(* Logix 5000 project; controller TFF vendor 1 type 14 code 107 rev 33.11; software revision 33.04 *)
// Mobius TFF

TASK HighPriority (periodic, rate 25 ms, priority 1, watchdog 2000 ms) : MainProgram   // High Priority Task
TASK MainTask (continuous, watchdog 500 ms) : Process, CCPSystem
TASK Task5ms (periodic, rate 5 ms, priority 10, watchdog 500 ms) : MainProgram5ms

MODULES
   Local : vendor 1 type 14 code 107 (Compact 0, rev 33.11)
      GATEWAY : ETHERNET-MODULE (Ethernet 10.20.60.222, rev 1.1, Output RPI 50 ms)
           GATEWAY:I   // Gateway data from hardware
           GATEWAY:O   // Gateway data from hardware
           GATEWAY:C   // Gateway data from hardware
      GWModbus : ETHERNET-MODULE (Ethernet 10.20.60.200, rev 1.1, Output RPI 50 ms)
           GWModbus:I.Data[56]   // R_PMC1 Unit
           GWModbus:I.Data[0]   // R_User Level
           GWModbus:I.Data[100]   // R_Warning Interface
           GWModbus:I.Data[101]   // R_Warning Interface
           GWModbus:I.Data[102]   // R_Warning Hardware
           GWModbus:I.Data[103]   // R_Warning Hardware
           GWModbus:I.Data[10]   // R_PMC1 Min limit
           GWModbus:I.Data[11]   // R_PMC1 Min limit
           GWModbus:I.Data[12]   // R_PMC1 Max limit
           GWModbus:I.Data[13]   // R_PMC1 Max limit
           GWModbus:I.Data[14]   // R_CalibStatus Status
           GWModbus:I.Data[15]   // R_CalibStatus Status
           GWModbus:I.Data[16]   // R_CalibStatus Unit
           GWModbus:I.Data[17]   // R_CalibStatus Unit
           GWModbus:I.Data[18]   // R_CalibStatus Value
           GWModbus:I.Data[19]   // R_CalibStatus Value
           GWModbus:I.Data[1]   // R_User Level
           GWModbus:I.Data[20]   // R_CalibLimits Offset Min
           GWModbus:I.Data[21]   // R_CalibLimits Offset Min
           GWModbus:I.Data[22]   // R_CalibLimits Offset Max
           GWModbus:I.Data[23]   // R_CalibLimits Offset Max
           GWModbus:I.Data[24]   // R_CalibLimits Slope Min
           GWModbus:I.Data[25]   // R_CalibLimits Slope Min
           GWModbus:I.Data[26]   // R_CalibLimits Slope Max
           GWModbus:I.Data[27]   // R_CalibLimits Slope Max
           GWModbus:I.Data[28]   // R_CalibValues Offset
           GWModbus:I.Data[29]   // R_CalibValues Offset
           GWModbus:I.Data[2]   // R_User N/A
           GWModbus:I.Data[30]   // R_CalibValues Slope
           GWModbus:I.Data[31]   // R_CalibValues Slope
           GWModbus:I.Data[32]   // R_CalibValues Temp
           GWModbus:I.Data[33]   // R_CalibValues Temp
           GWModbus:I.Data[34]   // R_CalibAct pH
           GWModbus:I.Data[35]   // R_CalibAct pH
           GWModbus:I.Data[36]   // R_CalibAct Elec
           GWModbus:I.Data[37]   // R_CalibAct Elec
           GWModbus:I.Data[38]   // R_CalibAct Temp
           GWModbus:I.Data[39]   // R_CalibAct Temp
           GWModbus:I.Data[3]   // R_User N/A
           GWModbus:I.Data[40]   // R_CalibAct NA
           GWModbus:I.Data[41]   // R_CalibAct NA
           GWModbus:I.Data[42]   // R_CalibTime Time
           GWModbus:I.Data[43]   // R_CalibTime Time
           GWModbus:I.Data[44]   // R_Warning Measurement
           GWModbus:I.Data[45]   // R_Warning Measurement
           GWModbus:I.Data[46]   // R_Warning Calibration
           GWModbus:I.Data[47]   // R_Warning Calibration
           GWModbus:I.Data[48]   // R_Warning Interface
           GWModbus:I.Data[49]   // R_Warning Interface
           GWModbus:I.Data[4]   // R_PMC1 Unit
           GWModbus:I.Data[50]   // R_Warning Hardware
           GWModbus:I.Data[51]   // R_Warning Hardware
           GWModbus:I.Data[52]   // R_User Level
           GWModbus:I.Data[53]   // R_User Level
           GWModbus:I.Data[54]   // R_User N/A
           GWModbus:I.Data[55]   // R_User N/A
           GWModbus:I.Data[57]   // R_PMC1 Unit
           GWModbus:I.Data[8]   // R_PMC1 Status
           GWModbus:I.Data[58]   // R_PMC1 Value
           GWModbus:I.Data[59]   // R_PMC1 Value
           GWModbus:I.Data[5]   // R_PMC1 Unit
           GWModbus:I.Data[60]   // R_PMC1 Status
           GWModbus:I.Data[61]   // R_PMC1 Status
           GWModbus:I.Data[62]   // R_PMC1 Min limit
           GWModbus:I.Data[63]   // R_PMC1 Min limit
           GWModbus:I.Data[64]   // R_PMC1 Max limit
           GWModbus:I.Data[65]   // R_PMC1 Max limit
           GWModbus:I.Data[66]   // R_CalibStatus Status
           GWModbus:I.Data[67]   // R_CalibStatus Status
           GWModbus:I.Data[68]   // R_CalibStatus Unit
           GWModbus:I.Data[69]   // R_CalibStatus Unit
           GWModbus:I.Data[6]   // R_PMC1 Value
           GWModbus:I.Data[70]   // R_CalibStatus Value
           GWModbus:I.Data[71]   // R_CalibStatus Value
           GWModbus:I.Data[72]   // R_CalibLimits Offset Min
           GWModbus:I.Data[73]   // R_CalibLimits Offset Min
           GWModbus:I.Data[74]   // R_CalibLimits Offset Max
           GWModbus:I.Data[75]   // R_CalibLimits Offset Max
           GWModbus:I.Data[76]   // R_CalibLimits Slope Min
           GWModbus:I.Data[77]   // R_CalibLimits Slope Min
           GWModbus:I.Data[78]   // R_CalibLimits Slope Max
           GWModbus:I.Data[79]   // R_CalibLimits Slope Max
           GWModbus:I.Data[7]   // R_PMC1 Value
           GWModbus:I.Data[80]   // R_CalibValues Offset
           GWModbus:I.Data[81]   // R_CalibValues Offset
           GWModbus:I.Data[82]   // R_CalibValues Slope
           GWModbus:I.Data[83]   // R_CalibValues Slope
           GWModbus:I.Data[84]   // R_CalibValues Temp
           GWModbus:I.Data[85]   // R_CalibValues Temp
           GWModbus:I.Data[86]   // R_CalibAct pH
           GWModbus:I.Data[87]   // R_CalibAct pH
           GWModbus:I.Data[88]   // R_CalibAct Elec
           GWModbus:I.Data[89]   // R_CalibAct Elec
           GWModbus:I.Data[9]   // R_PMC1 Status
           GWModbus:I.Data[90]   // R_CalibAct Temp
           GWModbus:I.Data[91]   // R_CalibAct Temp
           GWModbus:I.Data[92]   // R_CalibAct NA
           GWModbus:I.Data[93]   // R_CalibAct NA
           GWModbus:I.Data[94]   // R_CalibTime Time
           GWModbus:I.Data[95]   // R_CalibTime Time
           GWModbus:I.Data[96]   // R_Warning Measurement
           GWModbus:I.Data[97]   // R_Warning Measurement
           GWModbus:I.Data[98]   // R_Warning Calibration
           GWModbus:I.Data[99]   // R_Warning Calibration
           GWModbus:O.Data[12]   // W_CalibValue Temp
           GWModbus:O.Data[0]   // W_User Level
           GWModbus:O.Data[10]   // W_CalibValue Slope
           GWModbus:O.Data[11]   // W_CalibValue Slope
           GWModbus:O.Data[13]   // W_CalibValue Temp
           GWModbus:O.Data[24]   // W_SysTime Trigger
           GWModbus:O.Data[14]   // W_CalibProd Trigger
           GWModbus:O.Data[15]   // W_CalibProd Command
           GWModbus:O.Data[16]   // W_CalibProd Command
           GWModbus:O.Data[17]   // W_CalibProdVal Trigger
           GWModbus:O.Data[18]   // W_CalibProdVal Value
           GWModbus:O.Data[19]   // W_CalibProdVal Value
           GWModbus:O.Data[1]   // W_User Level
           GWModbus:O.Data[20]   // W_User Level
           GWModbus:O.Data[21]   // W_User Level
           GWModbus:O.Data[22]   // W_User Password
           GWModbus:O.Data[23]   // W_User Password
           GWModbus:O.Data[32]   // W_CalibValue Temp
           GWModbus:O.Data[25]   // W_SysTime Time
           GWModbus:O.Data[26]   // W_SysTime Time
           GWModbus:O.Data[27]   // W_CalibValue Trigger
           GWModbus:O.Data[28]   // W_CalibValue Offset
           GWModbus:O.Data[29]   // W_CalibValue Offset
           GWModbus:O.Data[2]   // W_User Password
           GWModbus:O.Data[30]   // W_CalibValue Slope
           GWModbus:O.Data[31]   // W_CalibValue Slope
           GWModbus:O.Data[33]   // W_CalibValue Temp
           GWModbus:O.Data[8]   // W_CalibValue Offset
           GWModbus:O.Data[34]   // W_CalibProd Trigger
           GWModbus:O.Data[35]   // W_CalibProd Command
           GWModbus:O.Data[36]   // W_CalibProd Command
           GWModbus:O.Data[37]   // W_CalibProdVal Trigger
           GWModbus:O.Data[38]   // W_CalibProdVal Value
           GWModbus:O.Data[39]   // W_CalibProdVal Value
           GWModbus:O.Data[3]   // W_User Password
           GWModbus:O.Data[4]   // W_SysTime Trigger
           GWModbus:O.Data[5]   // W_SysTime Time
           GWModbus:O.Data[6]   // W_SysTime Time
           GWModbus:O.Data[7]   // W_CalibValue Trigger
           GWModbus:O.Data[9]   // W_CalibValue Offset
      RACK_ACT350_WI101_200L : ETHERNET-MODULE (Ethernet 10.20.60.142, rev 1.1, Output RPI 50 ms)
      RACK_ACT350_WI101_500L : ETHERNET-MODULE (Ethernet 10.20.60.141, rev 1.1, Output RPI 50 ms)
      RACK_MURR_NODE0_SMART : ETHERNET-MODULE (Ethernet 10.20.60.131, rev 1.1, Output RPI 50 ms)
           RACK_MURR_NODE0_SMART:I   // Node 0 data from hardware
           RACK_MURR_NODE0_SMART:O.Data[0]   // MOM
           RACK_MURR_NODE0_SMART:O.Data[1]   // MOM
           RACK_MURR_NODE0_SMART:O.Data[2]   // MOM
           RACK_MURR_NODE0_SMART:O.Data[3]   // MOM
           RACK_MURR_NODE0_SMART:O.Data[4]   // MOM
           RACK_MURR_NODE0_SMART:O.Data[5]   // MOM
           RACK_MURR_NODE0_SMART:O.Data[6]   // Bus Control
           RACK_MURR_NODE0_SMART:O.Data[7]   // Bus Control
           RACK_MURR_NODE0_SMART:O   // Node 0 data from hardware
           RACK_MURR_NODE0_SMART:C   // Node 0 data from hardware
      RACK_MURR_NODE1_TFF20 : ETHERNET-MODULE (Ethernet 10.20.60.123, rev 1.1, Output RPI 5 ms)
           RACK_MURR_NODE1_TFF20:C   // Node 1 data from hardware
           RACK_MURR_NODE1_TFF20:I   // Node 1 data from hardware
           RACK_MURR_NODE1_TFF20:O   // Node 1 data from hardware
      RACK_MURR_NODE1_TFF40 : ETHERNET-MODULE (Ethernet 10.20.60.124, rev 1.1, Output RPI 5 ms)
           RACK_MURR_NODE1_TFF40:I   // Node 1 data from hardware
           RACK_MURR_NODE1_TFF40:O   // Node 1 data from hardware
           RACK_MURR_NODE1_TFF40:C   // Node 1 data from hardware
      RACK_MURR_NODE1_TFF80 : ETHERNET-MODULE (Ethernet 10.20.60.126, rev 1.1, Output RPI 5 ms)
           RACK_MURR_NODE1_TFF80:I   // Node 1 data from hardware
           RACK_MURR_NODE1_TFF80:O   // Node 1 data from hardware
           RACK_MURR_NODE1_TFF80:C   // Node 1 data from hardware
END_MODULES

TYPE AlarmAnalog :   // Analog Alarm UDT
STRUCT
   Override : BOOL;   // Alarm Override
   Disable : BOOL;   // Alarm Disabled
   LOLOAlarm : BOOL;   // LOLO Alarm Condition
   LOAlarm : BOOL;   // LO Alarm Condition
   HIAlarm : BOOL;   // HI Alarm Condition
   HIHIAlarm : BOOL;   // HIHI Alarm Condition
   LOLODisable : BOOL;   // LOLO Alarm Disable
   LODisable : BOOL;   // LO Alarm Disable
   HIDisable : BOOL;   // HI Alarm Disable
   HIHIDisable : BOOL;   // HIHI Alarm Disable
   LOLOAck : BOOL;   // LOLO Alarm Acknowledged
   LOAck : BOOL;   // LO Alarm Acknowledged
   HIAck : BOOL;   // HI Alarm Acknowledged
   HIHIAck : BOOL;   // HIHI Alarm Acknowledged
   HIHIEnable : BOOL;   // HIHI Alarm Always Enabled for Critical Safety Alarms
   FeedPumpEnable : BOOL;   // LOLO and LO Alarm conditionned on Feed Pump Enable
   TransferPumpEnable : BOOL;   // LOLO and LO Alarm conditionned on Transfer Pump Enable
   LOLOAlarmONS : BOOL;   // Saves last value of alarm
   LOAlarmONS : BOOL;   // Saves last value of alarm
   HIAlarmONS : BOOL;   // Saves last value of alarm
   HIHIAlarmONS : BOOL;   // Saves last value of alarm
   FeedPumpTag : DINT;   // Feed Pump Tag for Pump Enable function
   TransferPumpTag : DINT;   // Transfer Pump Tag for Pump Enable function
   Value : DINT;   // Alarm Value : 0= No Alarm. 1=Non-Critical. 2= Non-Critical Unacknowledged. 3=Critical. 4=Critical Unacknowledged.
   ValueHMI : DINT;   // Alarm Value for HMI: 0= No Alarm. 1=Non-Critical. 2= Non-Critical Unacknowledged. 3=Critical. 4=Critical Unacknowledged.
   LOLO : REAL;   // LOLO Alarm Set Point
   LO : REAL;   // LO Alarm Set Point
   HI : REAL;   // HI Alarm Set Point
   HIHI : REAL;   // HIHI Alarm Set Point
   PV : REAL;   // Process Variable Value
   LOLOTimer : TIMER;   // LOLO Alarm Timer
   LOLOTimerSP : DINT;   // LOLO Alarm Timer setpoint (sec)
   LOTimer : TIMER;   // LO Alarm Timer
   LOTimerSP : DINT;   // LO Alarm Timer setpoint (sec)
   HITimer : TIMER;   // HI Alarm Timer
   HITimerSP : DINT;   // HI Alarm Timer setpoint (sec)
   HIHITimer : TIMER;   // HIHI Alarm Timer
   HIHITimerSP : DINT;   // HIHI Alarm Timer setpoint (sec)
   EnableCfg : BOOL;   // Set to 1 to Configure \ Use Analog Alarm
END_STRUCT
END_TYPE

TYPE AlarmControl :   // Alarm Control UDT
STRUCT
   DESC : STRING25;   // Description
   EGU : STRING5;   // Unit
   InitAlarmconfig : BOOL;   // Initialize alarms config if the command is set from the HMI
   AlarmAck : BOOL;   // Alarm Acknowledge Flag
   AlarmHigh : BOOL;   // Critical Alarm Condition
   AlarmLow : BOOL;   // Non-Critical Alarm Condition
   AlarmHighUnack : BOOL;   // Critical Unacknowledged Alarm Condition
   AlarmLowUnack : BOOL;   // Non-Critical Unacknowledged Alarm Condition
   HighHMI : BOOL;   // Critical Alarm Condition (for HMI)
   LowHMI : BOOL;   // Non-Critical Alarm Condition (for HMI)
   HighUnackHMI : BOOL;   // Critical Unacknowledged Alarm Condition (for HMI)
   LowUnackHMI : BOOL;   // Non-Critical Unacknowledged Alarm Condition (for HMI)
   Horn : BOOL;   // Alarm Horn
   YellowLamp : BOOL;   // Non-Critical Alarm Indicator
   RedLamp : BOOL;   // Critical Alarm Indicator
   Current : BOOL;   // Current Alarm Status
   AckOutput : BOOL;   // Alarm Acknowledge Output
   FlashControl : BOOL;   // Flash Control
   LightingBannercfg : BOOL;   // Lighting Banner configuration (1= ON)
   EnableAllIn : BOOL;   // Enable All Alarms Input
   EnableAllOut : BOOL;   // Enable All Alarms Output
   DisableAllIn : BOOL;   // Disable All Alarms Input
   DisableAllOut : BOOL;   // Disable All Alarms Output
   NewAlarm : BOOL;   // True for 1 scan when new alarm is detected
   SilenceHorn : BOOL;   // Set true to Silence horn
   FlashTimer : TIMER;   // Flash Timer
   AckTimer : TIMER;   // Acknowledge Timer
   EnableAllTimer : TIMER;   // Enable All Alarms Timer
   DisableAllTimer : TIMER;   // Disable All Alarms Timer
   EnableAllAnaSigIn : BOOL;   // Enable All analog signal failure Alarms Input
   EnableAllAnaSigOut : BOOL;   // Enable All analog signal failure Alarms Output
   DisableAllAnaSigIn : BOOL;   // Disable All analog signal failure Alarms Input
   DisableAllAnaSigOut : BOOL;   // Disable All analog signal failure Alarms Output
   EnableAllAnaSigTimer : TIMER;   // Enable All analog signal failure Alarms Timer
   DisableAllAnaSigTimer : TIMER;   // Disable All analog signal failure Alarms Timer
   AlarmHighMem : BOOL;   // Critical Alarm Condition Mem
END_STRUCT
END_TYPE

TYPE AlarmDeviation :   // Deviation Alarm UDT
STRUCT
   Override : BOOL;   // Alarm Override
   Disable : BOOL;   // Alarm Disabled
   HIAlarm : BOOL;   // HI Deviation Alarm Condition
   HIHIAlarm : BOOL;   // HIHI Deviation Alarm Condition
   HIDisable : BOOL;   // HI Alarm Disable
   HIHIDisable : BOOL;   // HIHI Alarm Disable
   HIAck : BOOL;   // HI Alarm Acknowledged
   HIHIAck : BOOL;   // HIHI Alarm Acknowledged
   LOLOAlarmONS : BOOL;   // One shot when alarm occures
   HIAlarmONS : BOOL;   // One shot when alarm occures
   LOAlarmONS : BOOL;   // One shot when alarm occures
   HIHIAlarmONS : BOOL;   // One shot when alarm occures
   Value : DINT;   // Alarm Value
   ValueHMI : DINT;   // Alarm Value for HMI
   HI : REAL;   // HI Alarm Set Point
   HIHI : REAL;   // HIHI Alarm Set Point
   LOLOLim : REAL;   // LOLO Alarm Set Point (calculated)
   LOLim : REAL;   // LO Alarm Set Point (calculated)
   HILim : REAL;   // HI Alarm Set Point (calculated)
   HIHILim : REAL;   // HIHI Alarm Set Point (calculated)
   HITimer : TIMER;   // HI Alarm Timer
   HITimerSP : DINT;   // HI Alarm Timer setpoint (sec)
   HIHITimer : TIMER;   // HIHI Alarm Timer
   HIHITImerSP : DINT;   // HIHI Alarm Timer setpoint (sec)
   EnableCfg : BOOL;   // Set to enable alarm
END_STRUCT
END_TYPE

TYPE AnalogInput :   // Analog Input UDT
STRUCT
   TagName : STRING6;   // PID Tag Name
   TagDisplayName : STRING6;   // PID Tag Name
   OutofRange : BOOL;   // Out of Range
   FilterType : BOOL;   // Filter Type 0=LP, 1=Avg
   AveragingTotal : DINT;   // Averaging Filter Total
   Address : DINT;   // Input Address (RawAnalogInputArray)
   RawMin : DINT;   // Raw Minimum Range
   RawMax : DINT;   // Raw Maximum Range
   RawValue : DINT;   // Raw Value (Measuring value given by the I/O card)
   RawLowLimit : DINT;   // Raw Out of Range LO Limit
   RawHighLimit : DINT;   // Raw Out of Range HI Limit
   FilterUser : DINT;   // User Filter Value
   FilteredRaw : DINT;   // Raw Filtered Value
   FilterActual : REAL;   // Actual Filter Value
   ScaledMin : REAL;   // Scaled Minimum Range
   ScaledMax : REAL;   // Scaled Maximum Range
   CurrentValue : REAL;   // Current Value
   RangeMin : REAL;   // Scaled Minimum Range (Config Analog Points)
   RangeMax : REAL;   // Scaled Maximum Range (Config Analog Points)
   RangeMinSave : REAL;   // Scaled Minimum Range (previous)
   RangeMaxSave : REAL;   // Scaled Maximum Range (previous)
   RealCfg : BOOL;   // Set to 1 if real analog input is used. Set to 0 for soft input (derived data)
   EnableCfg : BOOL;   // Set to 1 to activate this Tag
   OverrideCfg : BOOL;   // Set to 1 to allow user to Overide alarm
   Desc : STRING25;   // Description
   EGU : STRING5;   // Unit
END_STRUCT
END_TYPE

TYPE AnalogOutput :   // Analog Output UDT
STRUCT
   Tag : STRING10;   // Tag name
   RawValue : DINT;   // Raw Value Send to I/O Card
   RawMin : DINT;   // Raw Min
   RawMax : DINT;   // Raw Max
   ScaledValue : REAL;   // Scaled Value
   ScaledMin : REAL;   // Scaled Minimum Range
   ScaledMax : REAL;   // Scaled Maximum Range
   EnableCfg : BOOL;   // Set to 1 to enable Analog Output
END_STRUCT
END_TYPE

TYPE ARC_pH :   // ARC pH Communication Structure
STRUCT
   SetCalibValues : BOOL;   // Set calibration values from HMI
   ActiveCalibration : BOOL;   // Current Active Calibration (0= Standrad, 1= Product)
   ActiveCalibrationSave : BOOL;   // Save state of Active Calibration
   AssignedCalibration : BOOL;   // Product Calibration is assigned
   ActiveInitial : BOOL;   // Initial Measurement of Product Calibration has been taken
   WarningSetCalib : BOOL;   // Verify/Set Calibration Data Warning from device
   ProductReadInitial : BOOL;   // Read command for the Product Calibration Initial Measurment
   ProductAssign : BOOL;   // Submit the Product Assign value command
   ProductAssignTime : DINT;   // Time of the last Product Assign
   ProductAssignONS : BOOL;   // ONS for Product Assignment
   R_CALIBSTATUS_Status : DINT;   // Calibration status from register 5318
   R_CALIBSTATUS_Unit : DINT;   // Calibration unit from register 5318
   R_CALIBSTATUS_Value : REAL;   // Calibration value from register 5318
   R_CALIBLIMITS_MinOffset : REAL;   // Calibration Minimum value for Offset from register 5480
   R_CALIBLIMITS_MaxOffset : REAL;   // Calibration Maximum value for Offset from register 5480
   R_CALIBLIMITS_MinSlope : REAL;   // Calibration Minimum value for Slope from register 5480
   R_CALIBLIMITS_MaxSlope : REAL;   // Calibration Maximum value for Slope from register 5480
   W_CALIBVALUES_Trigger : BOOL;   // Write to register 5448
   W_CALIBVALUES_Offset : REAL;   // Calibration offset to register 5448
   W_CALIBVALUES_Slope : REAL;   // Calibration slope to register 5448
   W_CALIBVALUES_Temp : REAL;   // Calibration temperature to register 5448
   R_CALIBVALUES_Offset : REAL;   // Calibration offset from register 5448
   R_CALIBVALUES_Slope : REAL;   // Calibration slope from register 5448
   R_CALIBVALUES_Temp : REAL;   // Calibration temperature from register 5448
   W_CALIBPROD_Trigger : BOOL;   // Write to register 5340
   W_CALIBPROD_Command : DINT;   // Product calibration command to register 5340
   W_CALIBPRODVAL_Trigger : BOOL;   // Write to register 5322
   W_CALIBPRODVAL_Value : REAL;   // Product calibration value to register 5322
   R_CALIBACTUAL_PH : REAL;   // pH at initial calibration from register 5560
   R_CALIBACTUAL_Voltage : REAL;   // Voltage at initial calibration from register 5560
   R_CALIBACTUAL_Temp : REAL;   // Temparature at initial calibration from register 5560
   R_CALIBACTUAL_NA : REAL;   // Unused from register 5560
   R_CALIBTIME_Time : DINT;   // Date Time of last calibration from register 5342 (UNIX)
   W_SYNCTIME_Trigger : BOOL;   // Write to register 8232
   W_SYNCTIME_Time : DINT;   // Time to register 8232 (UNIX)
   R_PMC1_Unit : DINT;   // Value unit from register 2090
   R_PMC1_Value : REAL;   // Value from register 2090
   R_PMC1_Status : DINT;   // Value Status from register 2090
   R_PMC1_Min : REAL;   // Value Minimum Limit from register 2090
   R_PMC1_Max : REAL;   // Value Maximum Limit from register 2090
   W_USER_Level : DINT;   // User Level to register 4288
   W_USER_Password : DINT;   // User Password to register 4288
   R_USER_Level : DINT;   // User Level from register 4288
   R_WARNING_Calib : DINT;   // Calibration warning from register 4736
END_STRUCT
END_TYPE

TYPE BagInflate :   // Inflate Bag
STRUCT
   cmd : BOOL;   // Command form HMI
   SP : REAL;   // Pressure Setpoint from HMI
   PV : REAL;   // Current Pressure
END_STRUCT
END_TYPE

TYPE CCPSystem :   // CCP System UDT
STRUCT
   Run : BOOL;   // Run Flag
   RunAuto : BOOL;   // Auto Run Flag
   Procedure : BOOL;   // Procedure Flag
   Complete : BOOL;   // Procedure Complete
   Download : BOOL;   // Manual Download
   Heartbeat : BOOL;   // CCPRuntime Heartbeat
   OperationDownloadFlag : BOOL;   // Legacy Tag. Not used by PLC
   OperationStartFlag : BOOL;   // Operation Start Flag
   Manual : BOOL;   // Recipe Pool Flag
   State : DINT;   // Machine State
   Language : DINT;   // Language Number
   ErrorPhase : DINT;   // Error in Phase #
   ErrorStep : DINT;   // Error in Step #
   Error : DINT;   // Error Description
   OperationNoInBatch : DINT;   // Legacy Tag. Not used by PLC
   EndPointer : DINT;   // End Operation Step Buffer Pointer
   Machine : STRING;   // Machine Name
   ProductID : STRING;   // Batch Product ID from Operation Header
   Description : STRING;   // Batch Description from Operation Header
   Created : STRING;   // Date and Time when the last operation has been downloaded in PLC
   Originator : STRING;   // Last saved by field from Operation Header
   Comment : STRING;   // Comment
   OperationName : STRING90;   // Name and path of last operation downloaded in PLC
   ConfigFile : STRING;   // Current configuration file used
   LastMod : STRING;   // Last Mod
   GradientBasis : STRING;   // Gradient Basis
   GradientVariable : STRING;   // Gradient Variable
   GradientSegments : STRING;   // Gradient Segments
   StateWatchDog : TIMER;   // If Downloading for longer than this time the state will reset to 0
   EventList : EventList;   // Event List Array
   BufferSteps : STRING25[251];   // Buffer Steps Array
   BufferEvents : STRING50[251];   // Buffer Events Array
   HETP_ON_OFF : BOOL;   // HETP (1 = Start , 0 = Stop)
   DefaultOnComplete : BOOL;   // At the end of recipe apply default flowpath (0 = Apply , 1 = Don't Apply)
END_STRUCT
END_TYPE

TYPE CCPSystem_Storage :
STRUCT
   Run : BOOL;   // Run Flag
   RunAuto : BOOL;   // Auto Run Flag
   Procedure : BOOL;   // Procedure Flag
   Complete : BOOL;   // Procedure Complete
   Download : BOOL;   // Manual Download
   Heartbeat : BOOL;   // CCPRuntime Heartbeat
   OperationDownloadFlag : BOOL;   // Legacy Tag. Not used by PLC
   OperationStartFlag : BOOL;   // Operation Start Flag
   TestAction : BOOL;   // Action Test Flag
   Manual : BOOL;   // Recipe Pool Flag
   State : DINT;   // Machine State
   Language : DINT;   // Language Number
   ErrorPhase : DINT;   // Error in Phase #
   ErrorStep : DINT;   // Error in Step #
   Error : DINT;   // Error Description
   OperationNoInBatch : DINT;   // Legacy Tag. Not used by PLC
   EndPointer : DINT;   // End Operation Step Buffer Pointer
   Machine : STRING;
   ProductID : STRING;
   Description : STRING;
   Created : STRING;
   Originator : STRING;
   Comment : STRING;
   OperationName : STRING90;
   ConfigFile : STRING;
   LastMod : STRING;
   GradientBasis : STRING;
   GradientVariable : STRING;
   GradientSegments : STRING;
   StateWatchDog : TIMER;   // If Downloading for longer than this time the state will reset to 0
END_STRUCT
END_TYPE

TYPE ChartMark :   // Chart Mark UDT
STRUCT
   In : BOOL;   // Chart Mark In
   Out : BOOL;   // Chart Mark Out
END_STRUCT
END_TYPE

TYPE Concentration :   // Concentration UDT
STRUCT
   VCF : REAL;   // Volume Concentration Factor
   CB : REAL;   // Protein Concentration
   Conc_Init : REAL;   // Initial Protein Concentration SP
   Conc_Final : REAL;   // Final Protein Concentration SP
   Conc_Final_Volume : REAL;   // Final Concentration Volume SP
   Final_Conc_Volume_Reached : BOOL;   // Final Concentration Volume Reached
   Final_Conc_Protein_Reached : BOOL;   // Final Protein Concentration Reached
   LogConcIn : BOOL;   // Log Concentration Input
   LogConcOut : BOOL;   // Log Concentration Output
   LogConcTimer : TIMER;   // Log Concentation Timer
END_STRUCT
END_TYPE

TYPE Configuration :   // Configuration UDT
STRUCT
   Reset : BOOL;   // Activate Reset Loop Configuration
   IndexA0 : DINT;   // Index AnalogOutput
   IndexAP : DINT;   // Index AnalogPoint
   IndexDP : DINT;   // Index DigitalPoint
   IndexDr : DINT;   // Index Drive
   IndeXValve : DINT;   // Index Valve
   IndexReset : DINT;   // Index Reset
   IndexCL : DINT;   // Index Control Loop
   IndexFlowpath : DINT;   // Index Flowpath
   IndexIOMod : DINT;   // Index IO Module
END_STRUCT
END_TYPE

TYPE ControlLoop :   // Control Loop UDT
STRUCT
   Tag : STRING5;   // Tag Name
   Desc : STRING25;   // Description
   LoopCfg : BOOL;   // Set to 1 to use this loop
   ManualEGU : STRING5;   // Unit of Manual Control Mode
   AutoEGU : STRING5;   // Unit of Auto Control Mode
   Auto1EGU : STRING5;   // Unit of Auto Control Mode 1
   Auto2EGU : STRING5;   // Unit of Auto Control Mode 2
   Auto3EGU : STRING5;   // Unit of Auto Control Mode 3
   Interlock : BOOL;   // Loop Interlock
   Enable : BOOL;   // Loop Enabled
   Manual : BOOL;   // Control Mode 0=Auto, 1=Manual
   Stable : BOOL;   // Loop Stable
   DBOK : BOOL;   // Control Within Deadband
   Status : INT;   // Status
   Auto1 : BOOL;   // Auto Control Mode 1
   Auto2 : BOOL;   // Auto Control Mode 2
   Auto3 : BOOL;   // Auto Control Mode 3
   Auto4 : BOOL;   // Auto Control Mode 4
   StepUp : BOOL;   // Increment CV
   StepDown : BOOL;   // Decrement CV
   RampEnable : BOOL;   // Ramp Enable
   RampUp : BOOL;   // Ramping UP
   RampDown : BOOL;   // Ramping Down
   RampStatus : BOOL;   // Ramping Status
   RampAutoOSR : BOOL;   // Auto Ramp One-Shot
   RampManualOSR : BOOL;   // Manual Ramp One-Shot
   PIDEnable : BOOL;   // PID Enabled
   ManualOSR : BOOL;   // Manual Mode One-Shot
   Auto1OSR : BOOL;   // Control Mode 1 One-Shot
   Auto2OSR : BOOL;   // Control Mode 2 One-Shot
   Auto3OSR : BOOL;   // Control Mode 3 One-Shot
   Auto4OSR : BOOL;   // Control Mode 4 One-Shot
   StepIncrement : DINT;   // Step Increment/Decrement Value
   CycleTime : DINT;   // Cycle Time (for modulating output)
   PV : REAL;   // Process Variable
   PVAuto1 : REAL;   // Process Variable for Control Mode Auto 1
   PVAuto2 : REAL;   // Process Variable for Control Mode Auto 2
   PVAuto3 : REAL;   // Process Variable for Control Mode Auto 3
   PVAuto4 : REAL;   // Process Variable for Control Mode Auto 4
   CV : REAL;   // Control Value
   SPAuto : REAL;   // Auto Set Point
   SPAutoSave : REAL;   // Auto Set Point (previous)
   SPAuto1 : REAL;   // Auto Set Point Mode 1
   SPAuto2 : REAL;   // Auto Set Point Mode 2
   SPAuto3 : REAL;   // Auto Set Point Mode 3
   SPAuto4 : REAL;   // Auto Set Point Mode 4
   SPManual : REAL;   // Manual Set Point
   SPManualSave : REAL;   // Manual Set Point (previous)
   RangeMin : REAL;   // Min EGU Range
   RangeMax : REAL;   // Max EGU Range
   SPRangeMin : REAL;   // Set Point Min EGU Range
   SPRangeMax : REAL;   // Set Point Max EGU Range
   RampRate : REAL;   // Ramp Rate
   RampRateSave : REAL;   // Ramp Rate (previous)
   RampStart : REAL;   // Ramp Start Value
   Deadband : REAL;   // Deadband
   DBLO : REAL;   // Low Deadband Value
   DBHI : REAL;   // High Deadband Value
   RampTimer : TIMER;   // Ramp Timer
   StableTimer : TIMER;   // Loop Stable Timer
   StableTime : DINT;   // Loop Stable Time setpoint (sec)
   PIDTimer : TIMER;   // PID Timer
   CycleTimer : TIMER;   // Cycle Timer (for modulating output)
   PID : PID;   // PID Instruction Data
   KP : REAL[3];   // Loop Gain from HMI
   KI : REAL[3];   // Loop Reset from HMI
   KD : REAL[3];   // Loop Rate from HMI
   DB : REAL[3];   // Loop Deadband from HMI
   On : BOOL;   // Turns all controll On
   DisOSR : BOOL;   // One Shot DisOSR
   OutputOn_OSR : BOOL;   // One Shot OutputOn_OSR
   OutputOff_OSR : BOOL;   // One Shot OutputOff_OSR
   DigitalOutput : BOOL;   // Output from loop in for descrete control
   RampCfg : BOOL;   // Set to 1 to Enable Ramp Option
   Auto1Cfg : BOOL;   // Set to 1 to use Auto 1 option
   Auto2Cfg : BOOL;   // Set to 1 to use Auto 2 option
   Auto3Cfg : BOOL;   // Set to 1 to use Auto 3 option
   Auto4Cfg : BOOL;   // Set to 1 to use Auto 4 option
   Auto1PVCfg : DINT;   // Set to Analog Point Number
   Auto2PVCfg : DINT;   // Set to Analog Point Number
   Auto3PVCfg : DINT;   // Set to Analog Point Number
   Auto4PVCfg : DINT;   // Set to Analog Point Number
   Auto1RangeMax : REAL;   // Set Point EGU Range Max
   Auto2RangeMax : REAL;   // Set Point EGU Range Max
   Auto3RangeMax : REAL;   // Set Point EGU Range Max
   Auto4RangeMax : REAL;   // Set Point EGU Range Max
   AutoSwitchEnable : BOOL;   // Set to 1 to allow loop to switch from auto1 to auto 2
   OutputAddress : INT;   // Set to analog output to use for this loop
   LoopStatus : INT;   // Loop Mode Status for HMI
END_STRUCT
END_TYPE

TYPE CriteriaFlag :   // Criteria Flag UDT
STRUCT
   Flag1 : BOOL;   // Criteria Flag 1 (1=ON , 0=OFF)
   Flag2 : BOOL;   // Criteria Flag 2 (1=ON , 0=OFF)
   Flag3 : BOOL;   // Criteria Flag 3 (1=ON , 0=OFF)
   Flag4 : BOOL;   // Criteria Flag 4 (1=ON , 0=OFF)
   Flag5 : BOOL;   // Criteria Flag 5 (1=ON , 0=OFF)
END_STRUCT
END_TYPE

TYPE CVTune :   // Control Valve Tuning Data Type
STRUCT
   ClosedRaw : REAL;   // Captured Raw Value When Valve is Closed
   OpenRaw : REAL;   // Captured Raw Value When Valve is Open
   MinOutput : REAL;   // Minimum output for tuning adjustment for valve
   MaxOutput : REAL;   // Maximum output for tuning adjustment for valve
   MinTimer : TIMER;   // Timer to capture closed raw value
   MaxTimer : TIMER;   // Timer to capture open raw value
   OSR : INT;   // One shot bits
   Activate : BOOL;   // Activate tuning function
   Enable : BOOL;   // Tuning routine is enabled
END_STRUCT
END_TYPE

TYPE DerivedData :   // DerivedData UDT
STRUCT
   HOLDUP : REAL;   // Holdup Volume
   FI101Q : REAL;   // Qmax Factor for FI101
   FI201Q : REAL;   // Qmax Factor for FI201
   FI401Q : REAL;   // Qmax Factor for FI401
   FI101K : REAL;   // K Factor for FI101
   FI201K : REAL;   // K Factor for FI201
   FI401K : REAL;   // K Factor for FI401
END_STRUCT
END_TYPE

TYPE Diafiltration :   // Diafiltration UDT
STRUCT
   Diaf_Volume : REAL;   // Diafiltration Volume
   Diaf_Init : REAL;   // Initial Diafiltration Volume SP
   Diaf_Final_Volume : REAL;   // Final Diafiltration Volume SP
   Snap : BOOL;   // Level Snapshot
   Final_Diaf_Volum_Reached : BOOL;   // Final Diafiltration Volume Reached
   Diaf_Snap_Value : REAL;   // Volume value snapped
   LogDiafIn : BOOL;   // Log Diafiltration Input
   LogDiafOut : BOOL;   // Log Diafiltration Output
   LogDiafTimer : TIMER;   // Log Diafiltration Timer
END_STRUCT
END_TYPE

TYPE DigitalPoint :   // Digital Point UDT
STRUCT
   Tag : STRING10;   // PID Tag to be Used for Display
   Desc : STRING25;   // Description to be Used for Display
   CurrentValue : BOOL;   // Current value of Tag
   AlarmCurrentValue : BOOL;   // Displays state of processed alarm input.
   AlarmAck : BOOL;   // Alarm Acknowledged
   Alarm : BOOL;   // Alarm
   Override : BOOL;   // Alarm Override
   Mimic : INT;   // Set color on HMI digital point mimic
   SoftInput : BOOL;   // Used as current value when RealInputCfg is set to 0
   Condition1 : BOOL;   // Enable Condition 1 Must be True to Enable alarm condition
   Condition2 : BOOL;   // Enable Condition 2 Must be True to Enable alarm condition
   Cond1Text : STRING;   // Condtion 1 Text
   Cond2Text : STRING;   // Condition 2 text
   DelayTimer : TIMER;   // Alarm Timer
   DelayTimerSP : DINT;   // Alarm Timer setpoint (sec)
   Priority : BOOL;   // Alarm Priority 0=Low, 1=High
   EnableCfg : BOOL;   // Set to True to configure point on system
   ActiveStateCFg : BOOL;   // Set to 0 to invert incomming state
   RealInputCfg : BOOL;   // Set to 1 to Use Hardwired Input. Set to 0 to disable Hardwired and use software condition
   InputAddressCfg : DINT;   // Set to address of hardwared input to be used on alarm
   AlarmCfg : BOOL;   // Set to 1 to Use alarm on this point
   AlarmStateCfg : BOOL;   // Set to 1 to alarm on a 0 to 1 transition. Set to zero to alarm on a 1 to 0 transition
   OverrideCfg : BOOL;   // set to 1 to allow user to Override alarm
   PriorityCfg : BOOL;   // Set to 1 to allow user to set Priority and Enable
   Cond1Cfg : BOOL;   // Set to 1 to Enable Condition
   Cond2Cfg : BOOL;   // Set to 1 to Enable Condition
   FlashingInputCfg : BOOL;   // Set to 1 for Heartbeat Style Inputs
   AlarmONS : BOOL;   // One shot when alarm occurs
END_STRUCT
END_TYPE

TYPE Drive :   // Pump Control UDT
STRUCT
   TagName : STRING10;   // Drive tag name
   Desc : STRING25;   // Drive Description
   Mode : BOOL;   // Control Mode
   ManualCommand : BOOL;   // Manual Command
   AutoCommand : BOOL;   // Auto Command
   RunCommand : BOOL;   // Run Command
   RunStatus : BOOL;   // Running Status
   RunInterlock : BOOL;   // Run Interlock
   RunInput : BOOL;   // Run Digital Input 0=No, 1=Yes
   OutputAddress : DINT;   // Run Command Output Address
   InputAddress : DINT;   // Running Input Address
   InterlockTimer : TIMER;   // Interlock Delay Timer
   RunOns : BOOL;   // Run one shot
   StopOns : BOOL;   // Stop One shot
   RunRequest : BOOL;   // Run request for auto or man mode
   Interlocked : BOOL;   // Drive is commanded to run but currently stopped by interlock
   EnableCfg : BOOL;   // Set to enable Drive
   ReverseCfg : BOOL;   // Set to enable reverse control
   Direction : BOOL;   // 0 = forward. 1 = reverse
   DirectionAddress : DINT;   // Direction Output Address
   DriveStatus : INT;   // Drive Status
   DriveLoopStatus : INT;   // Drive Loop Status
   DriveAlarmStatus : INT;   // Drive Alarm Status
   ValidFlowpath : BOOL;   // Valid flowpath flag
END_STRUCT
END_TYPE

TYPE EventList :
STRUCT
   Event : DINT[1000];   // Event List Array
   Value : REAL[1000];   // Value Array
   PreRunValue : REAL[1000];   // Pre Run Value
END_STRUCT
END_TYPE

TYPE Exchange_OUT :   // Exchange Output UDT
STRUCT
   AO01 : REAL;   // Exchange AO#1
   AO02 : REAL;   // Exchange AO#2
   AO03 : REAL;   // Exchange AO#3
   AO04 : REAL;   // Exchange AO#4
   DO01 : BOOL;   // Exchange DO#1
   DO02 : BOOL;   // Exchange DO#2
   DO03 : BOOL;   // Exchange DO#3
   DO04 : BOOL;   // Exchange DO#4
   DO05 : BOOL;   // Exchange DO#5
   DO06 : BOOL;   // Exchange DO#6
   DO07 : BOOL;   // Exchange DO#7
   DO08 : BOOL;   // Exchange DO#8
END_STRUCT
END_TYPE

TYPE FactorySettings :   // Factory Settings
STRUCT
   ProductName : STRING90;   // Product Name
   SerialNumber : STRING90;   // Serial Number
   ComputerName : STRING90;   // Computer Name
   ComputerDesc : STRING90;   // Computer Description
   DateFormat : STRING90;   // Date Format
   FlagUK : BOOL;   // Use UK Flag instead of US
   PCV101ClosedSP : REAL;   // PCV101 Closed SP
   PCV201ClosedSP : REAL;   // PCV201 Closed SP
   TCUDisableSP : REAL;   // TCU Disable SP
   BagInflateSP : REAL;   // Bag Inflate SP
END_STRUCT
END_TYPE

TYPE FaultRecordType :   // Fault Record Type UDT
STRUCT
   TimeLow : DINT;   // Lower 32 bits of the fault timestamp value
   TimeHigh : DINT;   // Upperer 32 bits of the fault timestamp value
   RecType : INT;   // Fault Type
   Code : INT;   // Unique code for the fault
   Info : DINT[8];   // Fault specific information
END_STRUCT
END_TYPE

TYPE FlowPath :   // Flow Path UDT
STRUCT
   Command : BOOL;   // Flow Path Command
   Status : BOOL;   // Flow Path Status
   Truth1 : DINT;   // Truth Table 1 (Valves 1-32)
   Truth2 : DINT;   // Truth Table 2 (Valves 33-64)
   Truth3 : DINT;   // Truth Table 3 (Valves 65-96)
   Truth4 : DINT;   // Truth Table 4 (Valves 97-128)
   Mask1 : DINT;   // Mask 1 (Valves 1-32)
   Mask2 : DINT;   // Mask 2 (Valves 33-64)
   Mask3 : DINT;   // Mask 3 (Valves 65-96)
   Mask4 : DINT;   // Mask 4 (Valves 97-128)
   Desc : STRING;   // Flow Path Description
END_STRUCT
END_TYPE

TYPE FlowPathControl :   // Flow Path Control UDT
STRUCT
   Flag : BOOL;   // Flow Path Command Flag
   Valve1 : DINT;   // Valve Control 1 (Valves 1-32)
   Valve2 : DINT;   // Valve Control 2 (Valves 33-64)
   Valve3 : DINT;   // Valve Control 3 (Valves 65-96)
   Valve4 : DINT;   // Valve Control 4 (Valves 97-128)
   MaxFlowPath : DINT;   // Maximum Number of Flow Paths
   Status : DINT;   // Flow Path Status
   StatusHMI : DINT;   // Flow Path Status for HMI
   Save : BOOL;   // Set to 1 to save Flowpath
   Restore : BOOL;   // Set to 1 to restore flowpath
   SaveOns : BOOL;   // one shot after save
   FlowpathEnable : BOOL[64];   // Enable Flowpath
   SaveStored : BOOL;   // Save the save cmd
   HoldOns : BOOL;   // one shot after hold
END_STRUCT
END_TYPE

TYPE FlowPathSetup :   // Flowpath Setup UDT
STRUCT
   Apply : BOOL;   // Apply Flow Path
   Number : DINT;   // Flow Path Number
   Prev : DINT;   // Previous Flow Path Number
   Mask_View : BOOL;   // View the Mask of selected Flowpath
   Mask_Save : BOOL;   // Save the Mask of selected Flowpath
   Truth_View : BOOL;   // View the Truth of selected Flowpath
   Truth_Save : BOOL;   // Save the Truth of selected Flowpath
   OpenAllValve : BOOL;   // Set the Flowpath 61 to Open All Valves
   CloseAllValve : BOOL;   // Set the Flowpath 62 to Close All Valves
END_STRUCT
END_TYPE

TYPE Gateway :   // Gateway UDT
STRUCT
   Inhibition : DINT;   // Inhibit \ Uninhibit Gateway Module
   Input : DINT[64];   // Swaped Data from Gateway
   Output : DINT[124];   // Swaped Data to Gateway
   RecipeAction_Digital : DINT[2];   // Data Send by PLC to Gateway (send from skid to customer) used as digital recipe action
   RecipeAction_Analog : REAL[20];   // Data Send by PLC to Gateway (send from skid to customer) used as analog recipe action
   RecipeCriteria_Digital : DINT[2];   // Data Read from the Gateway (receive from customer to skid) used as digital recipe criteria
   RecipeCriteria_Analog : REAL[20];   // Data Read from the Gateway (receive from customer to skid) used as analog recipe
   Watchdog_Heartbeat : BOOL;   // Gateway communication heartbeat
   Watchdog_Heartbeat_Timer : FBD_TIMER;   // Gateway communication heartbeat timer
   Watchdog_In_Ext : INT;   // Status data read by PLC (used to calculate customer watchdog)
   Watchdog_In_Skid : INT;   // Status data read by PLC (used to calculate skid watchdog)
   Watchdog_Out_Ext : INT;   // Status data send by PLC (used to calculate customer watchdog)
   Watchdog_Out_Skid : INT;   // Status data send by PLC (used to calculate skid watchdog)
   Index : DINT;   // Index
   Index2 : DINT;   // Index 2
END_STRUCT
END_TYPE

TYPE IO_Station :   // Station State UDT
STRUCT
   Node_Comm_Status_value : INT;   // Node Communication Status Value (get from status of hardware card)
   Node_Comm_Status : BOOL;   // Node Communication Status (0=Defect , 1=OK)
   Node_Internal_Defect_Status_value : INT;   // Node Internal Defect Status Value (at least one defect on the node : branch, slot, channel)
   Node_Internal_Defect_Status : BOOL;   // Node Internal Defect Status (0=Defect , 1=OK)
   Inhibition : DINT;   // Inhibit \ Uninhibit Station Module
   MOM_Mod_Config : BOOL[32];   // Activate \ Deactivate I/O Module (1 = Deactivate)
   MOM_Status : INT;   // Machine Option Management Status
   MOM_Restart : BOOL;   // 1 = Switch Off Voltage on modules , 0 = Restart the modules
   MOM_Enable_Config : BOOL;   // Enable modules configuration (avoid overwrite by options during the configuration)
END_STRUCT
END_TYPE

TYPE LinearGradient :   // Linear Gradient UDT
STRUCT
   Enable : BOOL;   // Linear Gradient Enable
   Hold : BOOL;   // Gradient Hold
   Segments : DINT;   // Number of Segments
   Variable : DINT;   // Gradient Variable (1=Time, 2=CVs, 3=Volume)
   Basis : DINT;   // Basis (1=Percent, 2=Conductivity)
   Segment : DINT;   // Current Segment
   State : DINT;   // Sets state of control : 0 = Disabled 1 = Running 2 = Paused
   Input : REAL;   // Input Value
   Result : REAL;   // Result
   X2 : REAL;   // Current Segment Duration
   Y1 : REAL;   // Current Start Value
   Y2 : REAL;   // Current End Value
   X : REAL[21];   // Gradient X Values (Durations)
   Y : REAL[21];   // Gradient Y Values (Set Points)
END_STRUCT
END_TYPE

TYPE LoggedValue :   // Logged Value UDT
STRUCT
   Value : REAL[8];   // Value to be logged in Audit Trail (used in Event section of configuration file)
END_STRUCT
END_TYPE

TYPE Membrane_Data :   // Membrane Data UDT
STRUCT
   Flux : REAL;   // Membrane Flux
   Area : REAL;   // Membrane Area SP
   Density : REAL;   // Density
   NWP_TCF : REAL;   // NWP Temperature correction factor
   NWP_TCF_Temp : INT;   // Temp. Temperature used in NWP calculation (INT)
   NWP_TCF_Lookup_25 : REAL[53];   // Lookup table for TCF
   AlarmStatus : INT;   // Alarm Status ( 0 = No Alarm , 1 = Non Critical Alarm , 2 = Critical Alarm )
END_STRUCT
END_TYPE

TYPE Memory_Data :   // This UDT is for putting the memory information returned by the Controller
STRUCT
   Reading_Request : BOOL;   // Request of Memory data reading
   Free_Mem_IO : DINT;   // Controler data: Free I/O Memory
   Free_Mem_DT : DINT;   // Controler data: Free Data & Logic Memory
   Free_Mem_Gen : DINT;   // Controler 1756-L55M16 only: Free Expansion Memory
   Free_Memory : DINT;   // Controler data: Total Free Memory (addition)
   Total_Mem_IO : DINT;   // Controler data: Total I/O Memory
   Total_Mem_DT : DINT;   // Controler data: Total Data & Logic Memory
   Total_Mem_Gen : DINT;   // Controler 1756-L55M16 only: Total Expansion Memory
   Total_Memory : DINT;   // Controler data: Total Memory (addition)
   Biggest_Gen_Mem_Size_Ava : DINT;   // Controler 1756-L55M16 only: Additionnal Expansion Memory
   Biggest_IO_Mem_Size_Ava : DINT;   // Controler 1756-L55M16 only: Largest contiguous block of Additionnal free Expansion Memory
   Biggest_DT_Mem_Size_Ava : DINT;   // Controler dsata: Largest contiguous block of Additionnal free Expansion Memory
   Total_Mem_DT_Real : REAL;   // Controler data: Total Data & Logic Memory
   Free_Mem_DT_Real : REAL;   // Controler data: Free Data & Logic Memory
   Used_Mem_DT_Real : REAL;   // Controler data: Used Data & Logic Memory
   Percentage_Used_DT : REAL;   // Controler data: Percentage of used Data & Logic Memory
END_STRUCT
END_TYPE

TYPE Mixer :
STRUCT
   Enable : BOOL;   // Enable Mixer Control Loop
   Mode : BOOL;   // Control Mode 0=Level, 1=Speed
   ModeONS : BOOL;   // Manual Mode One-Shot
   SPManual : REAL;   // Manual Speed Set Point
   SPAutoMin : REAL;   // Auto Max Speed Set Point
   SPAutoMax : REAL;   // Auto Min Speed Set Point
   LevelMin : REAL;   // Minimum Level
   LevelMax : REAL;   // Maximum Level
   CV : REAL;   // Control Value
   Alarm_Reset_Cmd : BOOL;   // Alarm Reset Command
   Alarm_Reset_Cmd_Timer : TIMER;   // Alarm Reset Command Timer
END_STRUCT
END_TYPE

TYPE OperatingTime :   // Operating Time Exceeded Control
STRUCT
   DayMax : REAL;   // Setpoint for Alarm Operating Time Exceeded
   HMICtrl : BOOL;   // Control Tag Reset on launch Workspace
   TimerCtrl : TIMER;   // Timer for set tag HMICtrl
   CountPre : DINT;   // Setpoint for Alarm in sec
   Counter : DINT;   // Second Counter for Alarm
END_STRUCT
END_TYPE

TYPE Operation :   // Operation UDT
STRUCT
   Step : DINT;   // Step Number
   Criteria1 : DINT;   // Criteria 1 Code
   Criteria1Operator : DINT;   // Criteria 1 Operator
   Boolean : DINT;   // Boolean
   Criteria2 : DINT;   // Criteria 2 Code
   Criteria2Operator : DINT;   // Criteria 2 Operator
   Action : DINT;   // Action Code
   Label : DINT;   // Label
   Criteria1Value : REAL;   // Criteria 1 Value
   Criteria2Value : REAL;   // Criteria 2 Value
   ActionValue : REAL;   // Action Value
END_STRUCT
END_TYPE

TYPE Options :   // Options UDT
STRUCT
   CCP_Report : BOOL;   // CCP Report
   InletFeed : BOOL;   // Feed Pump inlet
   InletFeed_Dis : BOOL;   // Feed Pump inlet Disabled
   FeedTank : BOOL;   // Feed Tank
   TransferFlow : BOOL;   // Transfer Flowmeter
   TankPH : BOOL;   // Tank pH Sensor
   TankCond : BOOL;   // Tank Conductivity Sensor
   FiltrateNoInstrum : BOOL;   // No Filtrate Instrument
   FiltrateNoInstrum_Dis : BOOL;   // No Filtrate Instrument Disabled
   FiltrateCondPH : BOOL;   // Filtrate Conductivity and PH
   FiltrateCondPHUV : BOOL;   // Filtrate Conductivity pH and UV
   FiltrateUltrasonicFlow : BOOL;   // Ultrasonic Filtrate Flowmeter instead of Magnetic
   FiltrateMagneticFlow : BOOL;   // Magnetic Filtrate Flowmeter instead of Ultrasonic
   SingleUsePH : BOOL;   // Single Use pH Sensor on Modbus Gateway
   External_IO : BOOL;   // External IO
   Gateway : BOOL;   // Gateway Anybus
   TFF80 : BOOL;   // TFF 80 Clamshell Installed
   TFF40 : BOOL;   // TFF 40 Clamshell Installed
   TFF20 : BOOL;   // TFF 20 Clamshell Installed
END_STRUCT
END_TYPE

TYPE PCV :
STRUCT
   SP : REAL;
   PV : REAL;
   ERREUR : REAL;
   CV : REAL;
   KP : REAL;
   KI : REAL;
   TP : REAL;
   TI : REAL;
   ACCU_TI : REAL;
   OpenRawValue : REAL;
   ClosedRawValue : REAL;
   RESET : BOOL;
END_STRUCT
END_TYPE

TYPE PCV_Calib :   // PCV Position Calibration
STRUCT
   Activate : BOOL;   // Calibration Command from HMI
   Enable : BOOL;   // PCV Calibration function enabled
   OSR : INT;   // One Shot bits
   Open_SP_Target : REAL;   // Open setpoint of PCV to achieve
   Close_SP_Target : REAL;   // Close setpoint of PCV to achieve
   Open_Timer : TIMER;   // Timer before save the raw value
   Close_Timer : TIMER;   // Timer before save the raw value
END_STRUCT
END_TYPE

TYPE PCV_Control :   // PCV Control UDT
STRUCT
   FullOpen : BOOL;   // fully open the valve without ramp
   FullOpenSP : REAL;   // target value of the valve opening
   FullOpenResetTimer : TIMER;   // Timer to reset full open command
   FullClose : BOOL;   // fully close the valve without ramp
   FullCloseSP : REAL;   // target value of the valve closing
   FullCloseResetTimer : TIMER;   // Timer to reset full close command
   ClosedStatusSP : REAL;   // Closed Status Setpoint
   ClosedStatus : BOOL;   // Closed Status
   CloseInterlocked : BOOL;   // Close Interlocked status for prohibit Manual Action on MHI
END_STRUCT
END_TYPE

TYPE Phases :   // Phase Control UDT
STRUCT
   Run : BOOL;   // Phase Run
   RunOSR : BOOL;   // Phase Run One-Shot
   Stop : BOOL;   // Phase Stop
   Hold : BOOL;   // Phase Hold
   Pause : BOOL;   // Phase Pause
   PauseOVR : BOOL;   // Pause Override
   Jump : BOOL;   // Phase Jump
   JumpPLC : BOOL;   // Phase Jump PLC
   Branch : BOOL;   // Branch Flag
   State : DINT;   // Phase State
   PendingStep : DINT;   // Pending Step Number
   JumpStep : DINT;   // Jump Step Number
   StartStep : DINT;   // Starting Step Number
   Crit1MetTime : DINT;   // Criteria 1 Met Timer
   NextStep : DINT;   // Next Step
   TotalSteps : DINT;   // Total Steps in Phase
   Label : DINT;   // Branch Label
   ActualStep : DINT;   // Actual Step
END_STRUCT
END_TYPE

TYPE PhaseTotalizer :   // Phase Totalizer UDT
STRUCT
   Enable : BOOL;   // Enable Totalizer
   PhaseEnable : BOOL;   // Enable Phase Totalizer
   StepEnable : BOOL;   // Enable Step Totalizer
   PauseEnable : BOOL;   // Enable Pause Totalizer
   UserEnable : BOOL;   // Enable User Totalizer
   ProcedureEnable : BOOL;   // Enable Procedure Totalizer
   PhaseReset : BOOL;   // Reset Phase Totalizer
   StepReset : BOOL;   // Reset Step Totalizer
   PauseReset : BOOL;   // Reset Pause Totalizer
   UserReset : BOOL;   // Reset User Totalizer
   PV : REAL;   // Totalizer Process Variable
   Phase : REAL;   // Phase Totalizer
   Step : REAL;   // Step Totalizer
   Pause : REAL;   // Pause Totalizer
   User : REAL;   // User Totalizer
   Procedure : REAL;   // Procedure Totalizer
   PVscale : REAL;   // PV Scaling
   PVsec : REAL;   // PV per second
   PVmin : REAL;   // PV Minimum Value
   Title : STRING10;   // Title to be displayed on status screen
   EGU : STRING10;   // EGU to display
   EnableCfg : BOOL;   // Set to one to use this totalizer
   SourceAddressCfg : INT;   // Enter analog Point # to be totalized
   SourceTypeCfg : BOOL;   // 0 For AnlogInput[] Source 1 For DerivedData.CVs Source
END_STRUCT
END_TYPE

TYPE PipeAnimation :   // Pipe Animation UDT
STRUCT
   PipeStat : BOOL[224];   // Pipe Animation Array
   PipeStatP1 : BOOL[224];   // Pipe Animation Array Line Pump 1
   PipeStatP2 : BOOL[224];   // Pipe Animation Array Line Pump 2
END_STRUCT
END_TYPE

TYPE Prompt :   // Prompt UDT
STRUCT
   Flag : BOOL;   // Flag
   PromptOK : BOOL;   // Type OK
   PromptYesNO : BOOL;   // Type Yes/No
   ResponseOK : BOOL;   // Input OK
   ResponseYes : BOOL;   // Input Yes
   ResponseNo : BOOL;   // Input No
   Pending : BOOL;   // Pending
   PromptONS : BOOL;   // One-Shot
   Step : DINT;   // Step Number
   Value : DINT;   // Value for PV+
END_STRUCT
END_TYPE

TYPE ScaleFiltering :   // Data for Scale Filtering
STRUCT
   CurrentFilter : INT;   // Type of filter used for Scale Filtering 0 = No Filtering 1 = Moving Average 2 = Exponential Linear Recursive
   Sample_Rate : DINT;   // Scale Filtering Sample Rate
   Timer : TIMER;   // Scale Filtering Timer
   WI101_Unfiltered : REAL;   // WI101 Unfiltered
   FeedBagVolume : REAL;   // Feed bag Volume based on WI101
   FeedBagVolume_Array : REAL[101];   // Array for Filter
   FeedBagVolume_MAVE : MOVING_AVERAGE;   // Feed Bag Volume Moving Average Filter structure
   WI201_Unfiltered : REAL;   // WI201 Unfiltered
   FiltrateVolume : REAL;   // Filtrate Volume based on WI201
   FiltrateVolume_Array : REAL[101];   // Array for Filter
   FiltrateVolume_MAVE : MOVING_AVERAGE;   // Filtrate Volume Moving Average Filter structure
   FiltrateVolume_MaveFiltered : REAL;   // Filtrate Volume value filtered by MAVE
   FiltrateVolume_ExpConst : REAL;   // Constant for Exponential Filter
   FiltrateVolume_ExpFiltered : REAL;   // Filtrate Volume value filtered by Exp
   Weight_ExpFiltered : REAL;   // Filtrate Weight filtered by Exp.
   Weight_MaveFiltered : REAL;   // Filtrate Weight filtered by MAVE
END_STRUCT
END_TYPE

TYPE STRING10 :   // 10 Character String
STRUCT
   LEN : DINT;
   DATA : SINT[10];
END_STRUCT
END_TYPE

TYPE STRING25 :   // 25 Character String
STRUCT
   LEN : DINT;
   DATA : SINT[26];
END_STRUCT
END_TYPE

TYPE STRING4 :   // 4 Character String
STRUCT
   LEN : DINT;
   DATA : SINT[4];
END_STRUCT
END_TYPE

TYPE STRING5 :   // 5 Character String
STRUCT
   LEN : DINT;
   DATA : SINT[5];
END_STRUCT
END_TYPE

TYPE STRING50 :   // 50 Character String
STRUCT
   LEN : DINT;
   DATA : SINT[50];
END_STRUCT
END_TYPE

TYPE STRING6 :   // 6 Character String
STRUCT
   LEN : DINT;
   DATA : SINT[6];
END_STRUCT
END_TYPE

TYPE STRING90 :   // 90 Character String
STRUCT
   LEN : DINT;
   DATA : SINT[90];
END_STRUCT
END_TYPE

TYPE SysControl :   // System Control Mode UDT
STRUCT
   DefaultIn : BOOL;   // Set System in Default In
   DefaultOut : BOOL;   // Set System in Default Out
   DefaultTimer : TIMER;   // Set System in Default Timer
   AllAutoIn : BOOL;   // Set System in All Auto In
   AllAutoOut : BOOL;   // Set System in All Auto Out
   AllAutoTimer : TIMER;   // Set System in All Auto Timer
   Simulate : BOOL;   // Enable Simulation Mode
   Simulate_Options : BOOL;   // Allow Options simulation
   Proc_Simulate : BOOL;   // Enable Process Simulation Mode
   Maintenance : BOOL;   // Enable Maintenance Mode
   DefaultStatus : BOOL;   // Default state status
   EnableSaveRestoreParam : BOOL;   // Enable save\restore parameters if condition are met
   UV_Auto_Zero_Cmd : BOOL;   // UV Auto Zero Command
   UV_Auto_Zero_Timer : TIMER;   // UV Auto Zero Timer
   Tare_WI101_Cmd : BOOL;   // Tank Weight Tare Command
   Tare_WI101_Timer : TIMER;   // Tank Weight Tare Timer
   ClearTare_WI101_Cmd : BOOL;   // Tank Weight Tare Clear Command
   ClearTare_WI101_Timer : TIMER;   // Tank Weight Tare Clear Timer
   Zero_WI101_Cmd : BOOL;   // Tank Weight Zero Command
   Zero_WI101_Timer : TIMER;   // Tank Weight Zero Timer
   Tare_PI001_Cmd : BOOL;   // Pressure PI001 Tare Command
   Tare_PI001_Timer : TIMER;   // Pressure PI001 Tare Timer
   Tare_PI101_Cmd : BOOL;   // Pressure PI101 Tare Command
   Tare_PI101_Timer : TIMER;   // Pressure PI101 Tare Timer
   Tare_PI201_Cmd : BOOL;   // Pressure PI201 Tare Command
   Tare_PI201_Timer : TIMER;   // Pressure PI201 Tare Timer
   Tare_PI401_Cmd : BOOL;   // Pressure PI401 Tare Command
   Tare_PI401_Timer : TIMER;   // Pressure PI401 Tare Timer
   Tare_PI601_Cmd : BOOL;   // Pressure PI601 Tare Command
   Tare_PI601_Timer : TIMER;   // Pressure PI601 Tare Timer
END_STRUCT
END_TYPE

TYPE SystemType :   // System Type UDT
STRUCT
   StatusTimer : TIMER;   // Evaluate Status Value Delay Timer
   Value : INT;   // Current value of system type (0-none, 1-chrom, 2-TFF)
   MoldType : INT;   // Current Value of the Installed Mold (123=TFF20, 124=TFF40, 126=TFF80)
   HMI_Value : INT;   // Current value of system mold from HMI (123=TFF20, 124=TFF40, 126=TFF80)
   PreviousValue : INT;   // Previous selected value; used to determine if new selection is made
   EnableSystemType : BOOL[32];   // Enable System Types
   CopyConfigFromMoldType0 : BOOL[32];   // Copy configuration data from Mold Type 0 to all other Mold Types
   CopyConfigFromMoldType1 : BOOL[32];   // Copy configuration data from Mold Type 1 to all other Mold Types
   CopyConfigFromMoldType2 : BOOL[32];   // Copy configuration data from Mold Type 2 to all other Mold Types
   CopyConfigFromMoldType3 : BOOL[32];   // Copy configuration data from Mold Type 3 to all other Mold Types
   CopyConfigFromMoldType4 : BOOL[32];   // Copy configuration data from Mold Type 4 to all other Mold Types
   DisableStatusCheck : BOOL;   // Disable Status Check; Allows for manual setting of System Type
   Initialize : BOOL;   // Upon new system selection, Initialize bit is set for any system Initialization required for setting up new system type
   Error : BOOL;   // Error bit if unable to determine system type
   ChangeCS : BOOL;   // Change CS Action from HMI
   NewCS : BOOL;   // New CS detected
   CopyParametersActive : BOOL;   // Manually set bit before setting Copy Configuration Data
   NewSystem_Timer : TIMER;   // One-Minute System change Timer
END_STRUCT
END_TYPE

TYPE TankManagement :   // UDT to Manage Tank
STRUCT
   Config : TankRange;   // Tank Range Configuration Management
   WeightConfiguration : TankRangeParameters[5];   // Tank Weight Range Parameters Management
   LevelConfiguration : TankRangeParameters[5];   // Tank Level Range Parameters Management
END_STRUCT
END_TYPE

TYPE TankRange :   // Update Tank Range Scaling & Alarming
STRUCT
   TankSelected : DINT;   // Tank Selected (0-None, 1-TK50, 2-TK100, 3-TK200, 4-TK500)
   TankSelectHMI : DINT;   // Tank Select HMI Use Only
   TankSelectPLC : DINT;   // Tank Select PLC
   Option_Current : DINT;   // Tank Current Option
   Option_Prev : DINT;   // Tank Previous Option
   Option_Simulate : DINT;   // Tank Option Simulated
   TMR : TIMER;
   ONS : DINT;   // One Shots
   MismatchAlarm : BOOL;   // Detects if Tank Selected is different from the actual connected tank
   Accept : BOOL;   // Operator Accepts Tank Selection
   ForceUpdate : BOOL;   // Force Tank Selection Update even if Tank Selection is same as Connected Tank
   Update : BOOL;   // Tank Selection Update Required
   UpdateComplete : BOOL;   // Tank Selection Update Complete
   WTUseDefault : BOOL;   // Load Default Alarm SP values
   LTUseDefault : BOOL;   // Load Default Alarm SP values
   Simulate : BOOL;   // Simulate Tank Option (0-Off, 1-On)
   AlarmStatus : INT;   // Alarm Status ( 0 = No Alarm , 1 = Non Critical Alarm , 2 = Critical Alarm )
   LevelHMI : REAL;   // Tank Level scaled for Tank animation in HMI
END_STRUCT
END_TYPE

TYPE TankRangeParameters :   // Update Tank Range Scaling & Alarming
STRUCT
   Desc : STRING25;   // Description
   ScaledMin : REAL;   // Scaled Min
   ScaledMin_PRE : REAL;   // Scaled Min Previous
   ScaledMax : REAL;   // Scaled Max
   ScaledMax_PRE : REAL;   // Scaled Max Previous
   RangeMin : REAL;   // Range Min
   RangeMin_PRE : REAL;   // Range Min Previous
   RangeMax : REAL;   // Range Max
   RangeMax_PRE : REAL;   // Range Max Previous
   Alm_LOLO : REAL;   // LOLO Alarm SP
   Alm_LOLO_PRE : REAL;   // LOLO Alarm SP Previous
   Alm_LO : REAL;   // LO Alarm SP
   Alm_LO_PRE : REAL;   // LO Alarm SP Previous
   Alm_HI : REAL;   // HI Alarm SP
   Alm_HI_PRE : REAL;   // HI Alarm SP Previous
   Alm_HIHI : REAL;   // HIHI Alarm SP
   Alm_HIHI_PRE : REAL;   // HIHI Alarm SP Previous
   Alm_LOLOTMR : DINT;   // LOLO Alarm Timer Preset
   Alm_LOLOTMR_PRE : DINT;   // LOLO Alarm Timer Preset Previous
   Alm_LOTMR : DINT;   // LO Alarm Timer Preset
   Alm_LOTMR_PRE : DINT;   // LO Alarm Timer Preset Previous
   Alm_HITMR : DINT;   // HI Alarm Timer Preset
   Alm_HITMR_PRE : DINT;   // HI Alarm Timer Preset Previous
   Alm_HIHITMR : DINT;   // HIHI Alarm Timer Preset
   Alm_HIHITMR_PRE : DINT;   // HIHI Alarm Timer Preset Previous
   Alm_Override : BOOL;   // Alarm Override
END_STRUCT
END_TYPE

TYPE TCUControl :   // TCU Control
STRUCT
   RunCommand : BOOL;   // Run Command
   ManualCommand : BOOL;   // Command Manual
   AutoCommand : BOOL;   // Command Auto
   Mode : BOOL;   // Control Mode (1= Manu)
   Interlock : BOOL;   // Interlock
   Interlocked : BOOL;   // Interlocked status for HMI
   SP_Disable : REAL;   // SP used when Disabled
   Offset : REAL;   // SP Offset when starting the TCU
   OffsetTimer : TIMER;   // Timer for active Offset
   OffsetTime : REAL;   // Timer for active Offset
   LevelMin : REAL;   // Level Minimum to start the TCU for Tank Temperature
   SPAutoSave : REAL;   // SP Auto Save for Offset ONS
   OffsetUp : BOOL;   // Offset direction to UP
   OffsetDown : BOOL;   // Offset direction to Down
END_STRUCT
END_TYPE

TYPE TimerControl :   // Timer Control UDT
STRUCT
   Tick : BOOL;   // 1 Second Tick to be used in HighPriority
   TickMainTask : BOOL;   // 1 Second Tick to be used in MainTask
   NewTickMainTask : BOOL;   // Flag to triger the main task Tick
   ResetAll : BOOL;   // Reset All Timers/Totalizers
   ResetProcedure : BOOL;   // Reset Procedure Timers/Totalizers
   Save : DINT;   // Saved Timer Value
   Seconds : DINT;   // Master Seconds Value
   Colon : STRING4;   // Colon ":"
   ColonZero : STRING4;   // Colon with Zero ":0"
   Cycle : DINT;   // Compute Value each 25ms (cycle time of HighPriority Task)
END_STRUCT
END_TYPE

TYPE Timers :   // Timers UDT
STRUCT
   Enable : BOOL;   // Enable Timer
   Reset : BOOL;   // Reset Timer
   TotalSeconds : REAL;   // Total Seconds Value
   Hours : DINT;   // HH Integer Value
   Minutes : DINT;   // MM Integer Value
   Seconds : DINT;   // SS Integer Value
   sHours : STRING4;   // HH String Value
   sMinutes : STRING4;   // MM String Value
   sSeconds : STRING4;   // SS String Value
   HMS : STRING25;   // HH:MM:SS Value
   LastHMS : STRING25;   // HH:MM:SS Value
END_STRUCT
END_TYPE

TYPE Totalizers :   // Totalizers UDT
STRUCT
   Enable : BOOL;   // Enable Totalizer
   Reset : BOOL;   // Reset Phase Totalizer
   PV : REAL;   // Totalizer Process Variable
   Total : REAL;   // Phase Totalizer
   PVscale : REAL;   // PV Scaling
   PVsec : REAL;   // PV per second
   PVmin : REAL;   // PV Minimum Value
   Title : STRING10;   // Title to be displayed on status screen
   LastTotal : REAL;   // a copy of the total at the last reset
   ResetTimer : TIMER;   // Reset timer for event log
   ResetONS : BOOL;   // Reset one-shot
END_STRUCT
END_TYPE

TYPE UserAlarm :   // User Alarm UDT
STRUCT
   NonCritical1 : BOOL;   // Set the User Non Critical Alarm 1
   Critical1 : BOOL;   // Set the User Critical Alarm 1
   NonCritical2 : BOOL;   // Set the User Non Critical Alarm 2
   Critical2 : BOOL;   // Set the User Critical Alarm 2
   SetUserAlarmC1ONS : BOOL;   // Set User Alarm 1 Oneshot
   SetUserAlarmC2ONS : BOOL;   // Set User Alarm 2 Oneshot
   SetUserAlarmNC1ONS : BOOL;   // Set User Alarm 1 Oneshot
   SetUserAlarmNC2ONS : BOOL;   // Set User Alarm 2 Oneshot
END_STRUCT
END_TYPE

TYPE UserTotalizerManagement :   // User Totalizer Management UDT
STRUCT
   LogUserIn : BOOL;   // Log User Totalizer Value
   LogUserOut : BOOL;   // Log User Totalizer Value
   StartUser : BOOL;   // Start User Totalizer
   ResetUserIn : BOOL;   // Reset User Totalizer
   ResetUserOut : BOOL;   // Reset User Totalizer
   LogUserTimer : TIMER;   // Log User Totalizer Timer
   ResetUserTimer : TIMER;   // Reset User Totalizer Timer
END_STRUCT
END_TYPE

TYPE Valve :   // Valve UDT
STRUCT
   Tag : STRING5;   // Tag Name
   Desc : STRING25;   // Description
   Control : BOOL;   // Valve Control
   Auto : BOOL;   // Auto Command
   Manual : BOOL;   // Manual Command (Force)
   Mode : BOOL;   // Control Mode
   ZSOpen : BOOL;   // Open Limit Switch
   ZSClose : BOOL;   // Closed Limit Switch
   ZSOpenEnable : BOOL;   // Enable Open Limit Switch
   ZSCloseEnable : BOOL;   // Enable Closed Limit Switch
   OpenStatus : BOOL;   // Open/On Status
   CloseStatus : BOOL;   // Closed/Off Status
   ZSOverride : BOOL;   // Limit Switch Override
   Priority : BOOL;   // Alarm Priority 0=Low, 1=High
   PriorityCfg : BOOL;   // Set to 1 to allow user to set Priority and Enable
   Alarm : BOOL;   // Alarm
   AlarmAck : BOOL;   // Alarm Acknowledged
   FailState : BOOL;   // Fail State 0=Closed, 1=Open
   Ports : BOOL;   // Number of Ports 0=2 way, 1=3 way
   OpenONS : BOOL;   // Open One-Shot
   CloseONS : BOOL;   // Close One-Shot
   EnableCfg : BOOL;   // Set to 1 to activate this Tag
   StatusWord : DINT;   // Valve Status word for HMI
   Status : DINT;   // Valve Status for Audit Trail
   ZSOpenAddress : DINT;   // Open Limit Switch Input Address
   ZSCloseAddress : DINT;   // Closed Limit Switch Input Address
   OutputAddress : DINT;   // Valve Output Address
   AlarmTimer : TIMER;   // Alarm Timer
   AlarmTimerSP : DINT;   // Alarm Timer setpoint (sec)
   AutoCloseTimer : TIMER;   // Auto Close Timer
   AlarmONS : BOOL;   // One shot when alarm occurs
   CloseInterlocked : BOOL;   // Close Interlocked status for prohibit Manual Action on MHI
END_STRUCT
END_TYPE
